(* IEC 61131-3 sources: codesys-framework/txt/application/WeVe Core (library)/60 Event, 4 files *)

(* ---- GeneralEvents.gvl.st ---- *)
VAR_GLOBAL CONSTANT

	cEv_Bookmark 								: DWORD := 16#00000000;

// [16#00000100 .. 16#000001FF] - Common
	cEv_PlcFirstCycleTask 						: UDINT := 16#00000100;
	cEv_MainPressureNotOk 						: UDINT := 16#00000101;

	cEv_ParameterUpdateRequest 					: UDINT := 16#00000102;
	cEv_ParameterUpdateNotAllowed 				: UDINT := 16#00000103;
	cEv_ParameterUpdateSucceeded 				: UDINT := 16#00000104;
	cEv_ParameterUpdateFailed 					: UDINT := 16#00000105;

	cEv_StartRequest 							: UDINT := 16#00000106;
	cEv_StopRequest 							: UDINT := 16#00000107;
	cEv_ResetRequest							: UDINT := 16#00000108;
	cEv_UserRequest								: UDINT := 16#00000109;
	cEv_StartRequestInvalid  					: UDINT := 16#0000010A;
	cEv_StopRequestInvalid  					: UDINT := 16#0000010B;
	cEv_ResetRequestInvalid  					: UDINT := 16#0000010C;
	cEv_UserRequestInvalid  					: UDINT := 16#0000010D;

	cEv_ModeRequest 							: UDINT := 16#0000010E;
	cEv_ModeRequestInvalid 						: UDINT := 16#0000010F;

// Module
	cEv_ModuleCommandTimeout 					: UDINT := 16#00000110;

// [16#00000200 - 16#000002FF] - Common	Safety
	cEv_SafetyNotOk 							: UDINT := 16#00000200;
	cEv_EmergencyStopActive 					: UDINT := 16#00000201;

END_VAR

(* ---- F_EventLevelToText.pou.st ---- *)
// Leesbare tekst voor een event-level, voor logregels.
FUNCTION F_EventLevelToText : STRING(20)
VAR_INPUT
	eLevel 			: E_EventLevels;
END_VAR
VAR
END_VAR

// --- BEGIN IMPLEMENTATION ---

CASE eLevel OF
	E_EventLevels.Success 						: F_EventLevelToText := 'Success';
	E_EventLevels.EventIsInformational 			: F_EventLevelToText := 'Info';
	E_EventLevels.EventIsWarning_NotUrgent 		: F_EventLevelToText := 'Warning';
	E_EventLevels.EventIsWarning_Urgent 		: F_EventLevelToText := 'Warning urgent';
	E_EventLevels.EventIsAlarm_OnlyLogLevel 	: F_EventLevelToText := 'Alarm log';
	E_EventLevels.EventIsAlarm_OperatorLevel 	: F_EventLevelToText := 'Alarm operator';
	E_EventLevels.EventIsAlarm_SupervisorLevel 	: F_EventLevelToText := 'Alarm supervisor';
ELSE
	F_EventLevelToText := 'Event';
END_CASE

(* ---- FB_Event.pou.st ---- *)
// Eén event: eenmalige melding (Log) of warning/alarm met toestand (Condition).
//
// Gebruik (via de EventGroup van de eigenaar):
//   - warning/alarm : elke cyclus Condition(xCondition := ..., scPayload := ...)
//   - eenmalig      : Log(scPayload := ...) bij het voorval
//   - reset         : Reset(), lukt enkel als de conditie weg is
//
// Boodschap: Config.sMessage met placeholders %0..%9, ingevuld met scPayload.asPayload[0..9].
// Logregel:  '<level> [<overgang>] | <id> | <subMachine>.<subMachineId> | <boodschap>'
//            bv. 'Alarm supervisor raised | 257 | 1.0 | Invalid air pressure'
// Tijdstempel en teller voegt de logger toe. Zonder logger houdt het event enkel zijn toestand bij.
FUNCTION_BLOCK FB_Event IMPLEMENTS I_Event
VAR_INPUT
END_VAR
VAR_OUTPUT
END_VAR
VAR
	_scConfig 		: SC_Event;
	_fbLogger 		: I_Logger;
	_xDisabled 		: BOOL;
	_xActive 		: BOOL;				// warning/alarm actief of gelatcht
	_xCondition 	: BOOL;				// conditie van de vorige aanroep, voor flankdetectie
	_scPayload 		: SC_EventPayload;	// payload van de laatste stijgende flank, voor cleared/reset
END_VAR

// --- BEGIN IMPLEMENTATION ---

(* ---- FB_EventGroup.pou.st ---- *)
// Basis voor de events van één eigenaar (mode, module of service).
//
// Een afgeleide groep levert:
//   - een enum per eigenaar, met Count als laatste element
//       E_AirPressureEvent : (PressureNok := 0, PressureLow, Count);
//   - de array van events
//       _afbEvents : ARRAY[0..E_AirPressureEvent.Count] OF FB_Event;   (slot Count blijft ongebruikt)
//   - GetEvent (met bounds check) en Count
//   - ConfigureEvents: één Configure-regel per event
//
// Wiring in FB_Application:
//   fbAirEvents : FB_AirPressureEvents(fbLogger := fbLogger, nSubMachine := 1, nSubMachineId := 0);
// Initialize() wordt eenmalig aangeroepen bij de opstart. Config wordt enkel dan gezet, nooit cyclisch.
FUNCTION_BLOCK ABSTRACT FB_EventGroup IMPLEMENTS I_EventGroup
VAR_INPUT
END_VAR
VAR_OUTPUT
END_VAR
VAR
	_fbLogger 			: I_Logger;
	_nSubMachine 		: USINT;
	_nSubMachineId 		: USINT;
	_xInitialized 		: BOOL;
END_VAR

// --- BEGIN IMPLEMENTATION ---
